TYPE TcoKukaKss_Status_v_9_3_x :
STRUCT
	ActionDescription : STRING(100);	
	State:TcoKukaKss_State_v_9_3_x;


END_STRUCT
END_TYPE

(* stored: Version 1.1.0.1, ProductVersion 3.1.4024.12
   DUT TcoKukaKss_Status_v_9_3_x: Id {eae09809-5c0e-496a-8147-5a37b8935664} *)
